Fanuc KAREL source: KO00046.KL

PROGRAM KO00046
%NOLOCKGROUP
%ENVIRONMENT MIR
VAR
  P1: POSITION
  P2: JOINTPOS
  F: BOOLEAN
  OUT: XYZWPR
BEGIN
  F = TRUE
  OUT = MIRROR(P1, P2, F)
END KO00046
